Yaskawa INFORM job: khoan10.JBI

/JOB
//NAME khoan10
//POS
///NPOS 22,0,0,0,0,0
///TOOL 9
///POSTYPE PULSE
///PULSE
C00000=-122907,48287,2678,-81935,-71000,-25622
C00001=-122907,52784,-1246,-82141,-71114,-23623
C00002=-122883,52870,-1083,-82149,-71101,-23635
C00003=-122895,52964,-905,-82143,-71106,-23648
C00004=-122938,53022,-796,-82127,-71127,-23656
C00005=-122993,53017,-806,-82108,-71153,-23656
C00006=-123032,52951,-931,-82095,-71172,-23647
C00007=-123039,52855,-1112,-82094,-71176,-23634
C00008=-123009,52774,-1265,-82106,-71163,-23623
C00009=-122957,52746,-1318,-82124,-71138,-23619
C00010=-122957,48247,2606,-81920,-71026,-25618
C00011=-133551,48468,3006,-78699,-76366,-25632
C00012=-133551,52957,-919,-78427,-76216,-23634
C00013=-133520,53037,-768,-78439,-76203,-23645
C00014=-133525,53134,-586,-78438,-76206,-23658
C00015=-133564,53201,-458,-78426,-76226,-23667
C00016=-133618,53208,-445,-78407,-76252,-23667
C00017=-133662,53152,-551,-78391,-76272,-23659
C00018=-133676,53058,-728,-78385,-76277,-23646
C00019=-133652,52971,-893,-78391,-76265,-23634
C00020=-133603,52931,-968,-78408,-76241,-23630
C00021=-133603,48441,2957,-78683,-76392,-25628
//INST
///DATE 2026/08/26 15:55
///COMM Generated using RoboDK
///ATTR SC,RW
///GROUP1 RB1
NOP
'Show Teknomotor QTC C4147-C-D
'B Spindle
MOVJ C00000 VJ=10.00 PL=1
MOVL C00001 V=200.0 PL=1
MOVL C00002 V=12.0 PL=1
MOVL C00003 V=12.0 PL=1
MOVL C00004 V=12.0 PL=1
MOVL C00005 V=12.0 PL=1
MOVL C00006 V=12.0 PL=1
MOVL C00007 V=12.0 PL=1
MOVL C00008 V=12.0 PL=1
MOVL C00009 V=12.0 PL=1
MOVL C00010 V=200.0 PL=1
MOVL C00011 V=200.0 PL=1
MOVL C00012 V=200.0 PL=1
MOVL C00013 V=12.0 PL=1
MOVL C00014 V=12.0 PL=1
MOVL C00015 V=12.0 PL=1
MOVL C00016 V=12.0 PL=1
MOVL C00017 V=12.0 PL=1
MOVL C00018 V=12.0 PL=1
MOVL C00019 V=12.0 PL=1
MOVL C00020 V=12.0 PL=1
MOVL C00021 V=200.0 PL=1
END
